// TIA Portal project "V20 Project_V20" (V20)

(* hardware
DEVICE "S7-1500/ET200MP station_1"  S7-1500 station
   slot 0: "Rail_0"  Rack  6ES7 590-1***0-0AA0
   slot 1: "PLC_2"  CPU 1515-2 PN  6ES7 515-2AM00-0AB0  V1.8
      slot 3: "CPU display_1"  6ES7591-1BA00-0AA0
      slot 32768: "PROFINET interface_1"  X1
         slot 32769: "Port_1"  X1 P1
         slot 32770: "Port_2"  X1 P2
      slot 33024: "PROFINET interface_2"  X2
         slot 33025: "Port_1"  X2 P1
*)

// ===== PLC "PLC_2"  CPU 1515-2 PN =====

FUNCTION_BLOCK "FB_CentreStand_Fix_Seq"   // FB1, STL
{ S7_Optimized_Access := 'TRUE' }
VERSION : 0.1
   VAR_INPUT
      iAutoRunning : Bool;
      iFixClamp : Bool;
      iFixEmpty : Bool;
      iFixTrayPresent : Bool;
      iFixUnclamp : Bool;
      iR1DropOver : Bool;
      iR1PickOver : Bool;
      iR2OperationOver : Bool;
      iR2ServiceActivated : Bool;
      iR2ServiceCompleted : Bool;
      iReset_fault : Bool;
      iRobotOutofZone : Bool;
      iSstMode : Bool;
      iSstPB : Bool;
   END_VAR
   VAR_OUTPUT
      qFixClamp : Bool;
      qFixUnclamp : Bool;
      qR1ReadytoDropTray : Bool;
      qR1ReadytoPickTray : Bool;
      qR2OperationStart : Bool;
   END_VAR
   VAR_IN_OUT
      iqR2ServiceActive : Bool;
      iqR2ServiceCompleted : Bool;
   END_VAR
   VAR
      StateNo : Int;
      s138_WaitBothRbtOutAl : Bool;
      s138_WaitBothRbtOutAl_T1 : Bool;
      s138_WaitBothRbtOutAl_T2 : Bool;
      s139_FixEmpty : Bool;
      s139_FixEmpty_T1 : Bool;
      s140_FixTrayPrsntRec : Bool;
      s140_FixTrayPrsntRec_T1 : Bool;
      s140_FixTrayPrsntRec_T2 : Bool;
      s141_FixUnclampCmd : Bool;
      s141_FixUnclampCmd_T1 : Bool;
      s142_TrayRdyDropFix : Bool;
      s142_TrayRdyDropFix_T1 : Bool;
      s143_RbtDropFixChkTr : Bool;
      s143_RbtDropFixChkTr_T1 : Bool;
      s144_RbtOutAreaDrop : Bool;
      s144_RbtOutAreaDrop_T1 : Bool;
      s145_FixClamp : Bool;
      s145_FixClamp_T1 : Bool;
      s146_Rbt2AlloyOpOver : Bool;
      s146_Rbt2AlloyOpOver_T1 : Bool;
      s147_FixUnclmpCmdOvr : Bool;
      s147_FixUnclmpCmdOvr_T1 : Bool;
      s148_RdyPickTrayWait : Bool;
      s148_RdyPickTrayWait_T1 : Bool;
      s149_RbtPickTrayChkEm : Bool;
      s149_RbtPickTrayChkEm_T1 : Bool;
      s191_WaitRbt2OutArea : Bool;
      s191_WaitRbt2OutArea_T1 : Bool;
      sSst : Bool;
      sSstPulse : Bool;
      sSstRise : Bool;
      sStWtResetRel : Bool;
      sStWtResetRel_T1 : Bool;
   END_VAR
   VAR_TEMP
      tOne : Bool;
   END_VAR
BEGIN

REGION Network 1
         O     #tOne;
         ON    #tOne;
         =     #tOne;
END_REGION

REGION Network 2: Create Single Step Pulse bit
         A     #iSstPB;
         FP    #sSstRise;
         =     #sSstPulse;
END_REGION

REGION Network 3: Create Single Step bit
         A     #iSstMode;
         A     #sSstPulse;
         ON    #iSstMode;
         =     #sSst;
END_REGION

REGION Network 4: Transition for STATE Num:0 Reset Released
         A     #sStWtResetRel;
         A     #iAutoRunning;
         =     #sStWtResetRel_T1;
END_REGION

REGION Network 5: STATE Num:0 Reset Released
         A(;
         O     #sStWtResetRel;
         ON    #iAutoRunning;
         );
         AN    #sStWtResetRel_T1;
         =     <??.?>;
         A     <??.?>;
         BLD   102;
         =     #sStWtResetRel;
         A     <??.?>;
         JNB   Label_0;
         L     0;
         T     #StateNo;
   Label_0:NOP   0;
END_REGION

REGION Network 6: Transition for STATE Num:138 Wait for Both Robots Out of Alloy Fixture Center Stand
         A     #s138_WaitBothRbtOutAl;
         AN    #sStWtResetRel;
         A     #sSst;
         =     <??.?>;
         A     <??.?>;
         A     #iRobotOutofZone;
         AN    #iFixTrayPresent;
         =     #s138_WaitBothRbtOutAl_T1;
         A     <??.?>;
         AN    #s138_WaitBothRbtOutAl_T1;
         A     #iRobotOutofZone;
         A     #iFixTrayPresent;
         =     #s138_WaitBothRbtOutAl_T2;
END_REGION

REGION Network 7: STATE Num:138 Wait for Both Robots Out of Alloy Fixture Center Stand
         A(;
         O     #s138_WaitBothRbtOutAl;
         O     #s149_RbtPickTrayChkEm_T1;
         O     #sStWtResetRel_T1;
         );
         AN    #sStWtResetRel;
         AN    #s138_WaitBothRbtOutAl_T1;
         AN    #s138_WaitBothRbtOutAl_T2;
         =     <??.?>;
         A     <??.?>;
         BLD   102;
         =     #s138_WaitBothRbtOutAl;
         A     <??.?>;
         JNB   Label_138;
         L     138;
         T     #StateNo;
   Label_138:NOP   0;
END_REGION

REGION Network 8: Transition for STATE Num:139 Fix Empty
         A     #s139_FixEmpty;
         AN    #sStWtResetRel;
         A     #sSst;
         A     #iFixEmpty;
         =     #s139_FixEmpty_T1;
END_REGION

REGION Network 9: STATE Num:139 Fix Empty
         A(;
         O     #s139_FixEmpty;
         O     #s138_WaitBothRbtOutAl_T1;
         );
         AN    #sStWtResetRel;
         AN    #s139_FixEmpty_T1;
         =     <??.?>;
         A     <??.?>;
         BLD   102;
         =     #s139_FixEmpty;
         A     <??.?>;
         JNB   Label_139;
         L     139;
         T     #StateNo;
   Label_139:NOP   0;
END_REGION

REGION Network 10: Transition for STATE Num:140 Fix Tray Present_Rec Operation pending
         A     #s140_FixTrayPrsntRec;
         AN    #sStWtResetRel;
         A     #sSst;
         =     <??.?>;
         A     <??.?>;
         A     #iFixTrayPresent;
         A     #iRobotOutofZone;
         AN    #iqR2ServiceCompleted;
         =     #s140_FixTrayPrsntRec_T1;
         A     <??.?>;
         AN    #s140_FixTrayPrsntRec_T1;
         A     #iFixTrayPresent;
         A     #iRobotOutofZone;
         A     #iqR2ServiceCompleted;
         =     #s140_FixTrayPrsntRec_T2;
END_REGION

REGION Network 11: STATE Num:140 Fix Tray Present_Rec Operation pending
         A(;
         O     #s140_FixTrayPrsntRec;
         O     #s138_WaitBothRbtOutAl_T2;
         );
         AN    #sStWtResetRel;
         AN    #s140_FixTrayPrsntRec_T1;
         AN    #s140_FixTrayPrsntRec_T2;
         =     <??.?>;
         A     <??.?>;
         BLD   102;
         =     #s140_FixTrayPrsntRec;
         A     <??.?>;
         JNB   Label_140;
         L     140;
         T     #StateNo;
   Label_140:NOP   0;
END_REGION

REGION Network 12: Transition for STATE Num:141 Fix Unclamp Cmd
         A     #s141_FixUnclampCmd;
         AN    #sStWtResetRel;
         A     #sSst;
         A     #iFixUnclamp;
         =     #s141_FixUnclampCmd_T1;
END_REGION

REGION Network 13: STATE Num:141 Fix Unclamp Cmd
         A(;
         O     #s141_FixUnclampCmd;
         O     #s139_FixEmpty_T1;
         );
         AN    #sStWtResetRel;
         AN    #s141_FixUnclampCmd_T1;
         =     <??.?>;
         A     <??.?>;
         BLD   102;
         =     #s141_FixUnclampCmd;
         A     <??.?>;
         JNB   Label_141;
         L     141;
         T     #StateNo;
   Label_141:NOP   0;
END_REGION

REGION Network 14: Actions for STATE Num:141 Fix Unclamp Cmd
         A     #s141_FixUnclampCmd;
         =     #qFixUnclamp;
END_REGION

REGION Network 15: Transition for STATE Num:142 Tray Rdy to Drop Fix- Wait for Robot Accept request
         A     #s142_TrayRdyDropFix;
         AN    #sStWtResetRel;
         A     #sSst;
         A     #iR1DropOver;
         =     #s142_TrayRdyDropFix_T1;
END_REGION

REGION Network 16: STATE Num:142 Tray Rdy to Drop Fix- Wait for Robot Accept request
         A(;
         O     #s142_TrayRdyDropFix;
         O     #s141_FixUnclampCmd_T1;
         );
         AN    #sStWtResetRel;
         AN    #s142_TrayRdyDropFix_T1;
         =     <??.?>;
         A     <??.?>;
         BLD   102;
         =     #s142_TrayRdyDropFix;
         A     <??.?>;
         JNB   Label_142;
         L     142;
         T     #StateNo;
   Label_142:NOP   0;
END_REGION

REGION Network 17: Actions for STATE Num:142 Tray Rdy to Drop Fix- Wait for Robot Accept request
         A     #s142_TrayRdyDropFix;
         =     #qR1ReadytoDropTray;
END_REGION

REGION Network 18: Transition for STATE Num:143 Robot Drop Fix and Check Tray Present
         A     #s143_RbtDropFixChkTr;
         AN    #sStWtResetRel;
         A     #sSst;
         A     #iFixTrayPresent;
         =     #s143_RbtDropFixChkTr_T1;
END_REGION

REGION Network 19: STATE Num:143 Robot Drop Fix and Check Tray Present
         A(;
         O     #s143_RbtDropFixChkTr;
         O     #s142_TrayRdyDropFix_T1;
         );
         AN    #sStWtResetRel;
         AN    #s143_RbtDropFixChkTr_T1;
         =     <??.?>;
         A     <??.?>;
         BLD   102;
         =     #s143_RbtDropFixChkTr;
         A     <??.?>;
         JNB   Label_143;
         L     143;
         T     #StateNo;
   Label_143:NOP   0;
END_REGION

REGION Network 20: Transition for STATE Num:144 Rbt Out of Area After Drop
         A     #s144_RbtOutAreaDrop;
         AN    #sStWtResetRel;
         A     #sSst;
         A     #iRobotOutofZone;
         =     #s144_RbtOutAreaDrop_T1;
END_REGION

REGION Network 21: STATE Num:144 Rbt Out of Area After Drop
         A(;
         O     #s144_RbtOutAreaDrop;
         O     #s143_RbtDropFixChkTr_T1;
         );
         AN    #sStWtResetRel;
         AN    #s144_RbtOutAreaDrop_T1;
         =     <??.?>;
         A     <??.?>;
         BLD   102;
         =     #s144_RbtOutAreaDrop;
         A     <??.?>;
         JNB   Label_144;
         L     144;
         T     #StateNo;
   Label_144:NOP   0;
END_REGION

REGION Network 22: Transition for STATE Num:145 Fix Clamp
         A     #s145_FixClamp;
         AN    #sStWtResetRel;
         A     #sSst;
         A     #iRobotOutofZone;
         A     #iFixClamp;
         =     #s145_FixClamp_T1;
END_REGION

REGION Network 23: STATE Num:145 Fix Clamp
         A(;
         O     #s145_FixClamp;
         O     #s140_FixTrayPrsntRec_T1;
         O     #s144_RbtOutAreaDrop_T1;
         );
         AN    #sStWtResetRel;
         AN    #s145_FixClamp_T1;
         =     <??.?>;
         A     <??.?>;
         BLD   102;
         =     #s145_FixClamp;
         A     <??.?>;
         JNB   Label_145;
         L     145;
         T     #StateNo;
   Label_145:NOP   0;
END_REGION

REGION Network 24: Actions for STATE Num:145 Fix Clamp
         A     #s145_FixClamp;
         =     #qFixClamp;
END_REGION

REGION Network 25: Transition for STATE Num:146 Robot-2 All Alloys Pick Or Drop Operation over
         A     #s146_Rbt2AlloyOpOver;
         AN    #sStWtResetRel;
         A     #sSst;
         A     #iR2OperationOver;
         =     #s146_Rbt2AlloyOpOver_T1;
END_REGION

REGION Network 26: STATE Num:146 Robot-2 All Alloys Pick Or Drop Operation over
         A(;
         O     #s146_Rbt2AlloyOpOver;
         O     #s145_FixClamp_T1;
         );
         AN    #sStWtResetRel;
         AN    #s146_Rbt2AlloyOpOver_T1;
         =     <??.?>;
         A     <??.?>;
         BLD   102;
         =     #s146_Rbt2AlloyOpOver;
         A     <??.?>;
         JNB   Label_146;
         L     146;
         T     #StateNo;
   Label_146:NOP   0;
END_REGION

REGION Network 27: Actions for STATE Num:146 Robot-2 All Alloys Pick Or Drop Operation over
         A     #s146_Rbt2AlloyOpOver;
         =     #qR2OperationStart;
         A     #iR2ServiceActivated;
         S     #iqR2ServiceActive;
         A     #iR2OperationOver;
         A     #iqR2ServiceActive;
         R     #iqR2ServiceActive;
END_REGION

REGION Network 28: Transition for STATE Num:147 Fix Unclamp Cmd After Opern over
         A     #s147_FixUnclmpCmdOvr;
         AN    #sStWtResetRel;
         A     #sSst;
         A     #iFixUnclamp;
         =     #s147_FixUnclmpCmdOvr_T1;
END_REGION

REGION Network 29: STATE Num:147 Fix Unclamp Cmd After Opern over
         A(;
         O     #s147_FixUnclmpCmdOvr;
         O     #s140_FixTrayPrsntRec_T2;
         O     #s191_WaitRbt2OutArea_T1;
         );
         AN    #sStWtResetRel;
         AN    #s147_FixUnclmpCmdOvr_T1;
         =     <??.?>;
         A     <??.?>;
         BLD   102;
         =     #s147_FixUnclmpCmdOvr;
         A     <??.?>;
         JNB   Label_147;
         L     147;
         T     #StateNo;
   Label_147:NOP   0;
END_REGION

REGION Network 30: Actions for STATE Num:147 Fix Unclamp Cmd After Opern over
         A     #s147_FixUnclmpCmdOvr;
         =     #qFixUnclamp;
END_REGION

REGION Network 31: Transition for STATE Num:148 Rdy to Pick Tray After Oprn Over- Wait for Robot Accept Request
         A     #s148_RdyPickTrayWait;
         AN    #sStWtResetRel;
         A     #sSst;
         A     #iR1PickOver;
         =     #s148_RdyPickTrayWait_T1;
END_REGION

REGION Network 32: STATE Num:148 Rdy to Pick Tray After Oprn Over- Wait for Robot Accept Request
         A(;
         O     #s148_RdyPickTrayWait;
         O     #s147_FixUnclmpCmdOvr_T1;
         );
         AN    #sStWtResetRel;
         AN    #s148_RdyPickTrayWait_T1;
         =     <??.?>;
         A     <??.?>;
         BLD   102;
         =     #s148_RdyPickTrayWait;
         A     <??.?>;
         JNB   Label_148;
         L     148;
         T     #StateNo;
   Label_148:NOP   0;
END_REGION

REGION Network 33: Actions for STATE Num:148 Rdy to Pick Tray After Oprn Over- Wait for Robot Accept Request
         A     #s148_RdyPickTrayWait;
         =     #qR1ReadytoPickTray;
         A     #iR1PickOver;
         R     #iqR2ServiceCompleted;
END_REGION

REGION Network 34: Transition for STATE Num:149 Robot Picked Tray and Check Tray Loc Empty
         A     #s149_RbtPickTrayChkEm;
         AN    #sStWtResetRel;
         A     #sSst;
         A     #iFixEmpty;
         =     #s149_RbtPickTrayChkEm_T1;
END_REGION

REGION Network 35: STATE Num:149 Robot Picked Tray and Check Tray Loc Empty
         A(;
         O     #s149_RbtPickTrayChkEm;
         O     #s148_RdyPickTrayWait_T1;
         );
         AN    #sStWtResetRel;
         AN    #s149_RbtPickTrayChkEm_T1;
         =     <??.?>;
         A     <??.?>;
         BLD   102;
         =     #s149_RbtPickTrayChkEm;
         A     <??.?>;
         JNB   Label_149;
         L     149;
         T     #StateNo;
   Label_149:NOP   0;
END_REGION

REGION Network 36: Actions for STATE Num:149 Robot Picked Tray and Check Tray Loc Empty
         A     #s149_RbtPickTrayChkEm;
         R     #iqR2ServiceCompleted;
END_REGION

REGION Network 37: Transition for STATE Num:191 Wait For Robot-2 Out Of Area
         A     #s191_WaitRbt2OutArea;
         AN    #sStWtResetRel;
         A     #sSst;
         A     #iRobotOutofZone;
         =     #s191_WaitRbt2OutArea_T1;
END_REGION

REGION Network 38: STATE Num:191 Wait For Robot-2 Out Of Area
         A(;
         O     #s191_WaitRbt2OutArea;
         O     #s146_Rbt2AlloyOpOver_T1;
         );
         AN    #sStWtResetRel;
         AN    #s191_WaitRbt2OutArea_T1;
         =     <??.?>;
         A     <??.?>;
         BLD   102;
         =     #s191_WaitRbt2OutArea;
         A     <??.?>;
         JNB   Label_191;
         L     191;
         T     #StateNo;
   Label_191:NOP   0;
END_REGION
END_FUNCTION_BLOCK

FUNCTION_BLOCK "Block_1"   // FB1, LAD
{ S7_Optimized_Access := 'TRUE' }
BEGIN

REGION Network 1
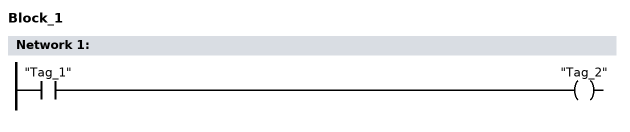
   RUNG wire#powerrail
      Contact( "Tag_1" )
      Coil( "Tag_2" )
   END_RUNG
   // the same network as SCL:
   "Tag_2" := "Tag_1";
END_REGION
END_FUNCTION_BLOCK

ORGANIZATION_BLOCK "Main"   // OB1, LAD, ProgramCycle
TITLE = "Main Program Sweep (Cycle)"
{ S7_Optimized_Access := 'TRUE' }
VERSION : 0.1
   VAR_INPUT
      Initial_Call : Bool;   // Initial call of this OB
      Remanence : Bool;   // =True, if remanent data are available
   END_VAR
BEGIN
END_ORGANIZATION_BLOCK

// ===== library types =====

// folder: SM-Modules

FUNCTION_BLOCK "PR_TT3PosControl"   // FB335, LAD
TITLE = PR_TT3PosControl
{ S7_Optimized_Access := 'TRUE' }
AUTHOR : Virendra Sharma
FAMILY : Wipro_Pari
NAME : SM0106022020
VERSION : 0.1
   VAR_INPUT
      iResetFaults : Bool;   // Reset Fault input
      iControlOn : Bool;   // Control On Input
      iPos1Cmd : Bool;   // Zero degree position command (Home position)
      iPos2Cmd : Bool;   // Plus 90 degree position command
      iPos3Cmd : Bool;   // Minus 90 degree position command
      iPos1StopSens : Bool;   // zero degree position stop sensor
      iPos2StopSens : Bool;   // Plus 90 degree position stop sensor
      iPos3StopSens : Bool;   // Minus 90 degree position stop sensor
      iTimeForPosOver : Time;   // Timer Value for position over
      iTimeForVFDStop : Time;   // Time value for VFD stop
      iPositiveOTLS : Bool;   // Positive direction over travel limit swithch
      iNegativeOTLS : Bool;   // Negative direction over travel limit swithch
      iFwdInterlock : Bool;   // Connect Forward Interlock Conditions
      iRevInterlock : Bool;   // Connect Reverse Interlock Conditions
      iVFDRunning : Bool;
   END_VAR
   VAR_OUTPUT
      qPos1Over : Bool;   // Zero position over
      qPos2Over : Bool;   // Plus 90 position
      qPos3Over : Bool;   // Minus 90 position over
      qVFDFwd : Bool;   // VFD Rotating Forward
      qVFDRev : Bool;   // VFD Rotating Reverse
      qModuleFault : Bool;   // Error Module Fault
      qError : Array[0..7] of Bool;   // Error Forward Interlock
      qMsg : Array[0..7] of Bool;
   END_VAR
   VAR
      sFaultReset : Bool;
      sFwdCmdOn : Bool;
      sDriveRdyFrCmd : Bool;
      sTimeForPosOver : Time;
      sTimeForVFDStop : Time;
      sRevCmdOn : Bool;
      sCtrlFrmNet : Bool;
      sRefFrmNet : Bool;
      sTimerOn : Bool;
      s0PosCmdActive : Bool;
      s0PosActiveForFwd : Bool;
      s0PosActiveForRev : Bool;
      s0PosActiveForFwdOver : Bool;
      s0PosActiveForRevOver : Bool;
      s0PosOverTON : TON_TIME;
      sMinus90PosActiveForRev : Bool;
      sMinus90PosCmdActive : Bool;
      sMinus90PosOverTON : TON_TIME;
      sMinus90PosActiveForFwdOver : Bool;
      sMinus90PosActiveForRevOver : Bool;
      sPlus90PosActiveForFwd : Bool;
      sPlus90PosCmdActive : Bool;
      sPlus90PosOverTON : TON_TIME;
      sPlus90PosActiveForFwdOver : Bool;
      sPlus90PosActiveForRevOver : Bool;
      sTTAtPos0 : Bool;
      sTTAtPos0Done : Bool;
      sTTAtPosMinus90 : Bool;
      sTTAtPosMinus90Done : Bool;
      sTTAtPosPlus90 : Bool;
      sTTAtPosPlus90Done : Bool;
      sPuls : Array[0..16] of Bool;
   END_VAR
   VAR RETAIN
      sTargetPos : Word;
      sLastPos : Word;
   END_VAR
   VAR
      sVFDFwdRunning : Bool;
      sVFDRunningDlyDn : TON_TIME;
      sVFDRevRunning : Bool;
      sFwdInterlockErr : Bool;
      sRevInterlockErr : Bool;
      sPositiveOTLSErr : Bool;
      sNegativeOTLSErr : Bool;
      sVFDStopped : Bool;
   END_VAR
   VAR RETAIN
      sFwdActiveFor1ToPos2 : Bool;
      sRevAvtiveFor1ToPos3 : Bool;
      sFwdActiveFor3ToPos1 : Bool;
      sRevAvtiveFor2ToPos1 : Bool;
   END_VAR
   VAR_TEMP   // added for the SCL form of the ladder/FBD networks
      _w1 : Bool;
      _w2 : Bool;
      _w3 : Bool;
      _w4 : Bool;
      _w5 : Bool;
      _w6 : Bool;
   END_VAR
   // // qError[1] : Error Reverse Interlock
   // // qError[2] : Error Forward Interlock
   // // qError[3] : Turn Table over traveled at positive side
   // // qError[4] : Turn Table over traveled at negative side
   // // qError[0] : Error VFD Stopped
   // // qMsg[0] : TT not referenced.
BEGIN

REGION Network 1: Header
   // ==============================================================================
   //  Company: Precision Automation & Robotics India Ltd. (WIPRO-PARI)
   // ------------------------------------------------------------------------------
   //  Item Code: SM0106022020
   //  Author/Created by: Virendra Sharma
   //  Reviewed/Checked by: Sandip Chavanke
   //  First Release on: 11-Oct-2023
   //  Latest update on: 11-Oct-2023
   // ------------------------------------------------------------------------------
   //  Tested with: CPU firmware, model or simulator testing
   //  Engineering/Editor: TIA Portal V17
   // ------------------------------------------------------------------------------
   //  Restrictions: More then 3 Position of turn table
   //  Dependencies/Requirements:
   //  <hardware, technology package, memory needed, data types (UDT's), other blocks, etc.>
   // ------------------------------------------------------------------------------
   //  Change Log:
   //  Ver.	Date		Changed by		Details of changes
   //  1.0	11-10-2023	Virendra Sharma 	First release version- 1.0
   // ------------------------------------------------------------------------------
   //  Functionality: This Module is to control the motion of VFD that controls Turn Table with 3 distinctive positions,
   //  like home or Path1 (0 Degree), Path3 (Minus 90 Degree), and path2 (Plus 90 Degree) positions.
   //  Each position is provided with a 'position sensor' to confirm the position of the Turn Table and to stop the Turn Table at the given position.
   //  The position of the turn table is defined by where the main stopper is located.
   //  <include block inputs, outputs, in-outs>
   //  Inputs
   //  1. iResetFaults : Bool
   //  2. iControlOn : Bool
   //  3. iPos1Cmd : Bool
   //  4. iPos2Cmd : Bool
   //  5. iPos3Cmd : Bool
   //  6. iPos1StopSens : Bool
   //  7. iPos2StopSens : Bool
   //  8. iPos3StopSens : Bool
   //  9. iTimeForPosOver : Time
   //  10. iTimeForVFDStop : Time
   //  11. iPositiveOTLS : Bool
   //  12. iNegativeOTLS : Bool
   //  13. iFwdInterlock : Bool
   //  14. iRevInterlock : Bool
   // 
   //  Outputs
   //  1. qPos1Over : Bool
   //  2. qPos2Over : Bool
   //  3. qPos3Over : Bool
   //  4. qVFDFwd : Bool
   //  5. qVFDRev : Bool
   //  6. qModuleFault : bool
   //  7. qError : Array [0..31] of Bool
   //  8. qMsg : Array [0..31] of Bool  
   // 
   //  In-outs
   //  NA
   // ------------------------------------------------------------------------------
   //  Errors reported:
   //  1. Error 0 : Error VFD Stopped
   //  2. Error 1 : Error Reverse Interlock 
   //  3. Error 2 : Error Forward Interlock 
   //  4. Error 3 : Turn Table over traveled at positive side
   //  5. Error 4 : Turn Table over traveled at negative side
   //  Messages reported:
   //  1. Message 0 : TT not referenced.
   // ==============================================================================
END_REGION

REGION Network 2: Fault Reset
   // Error reset request flag
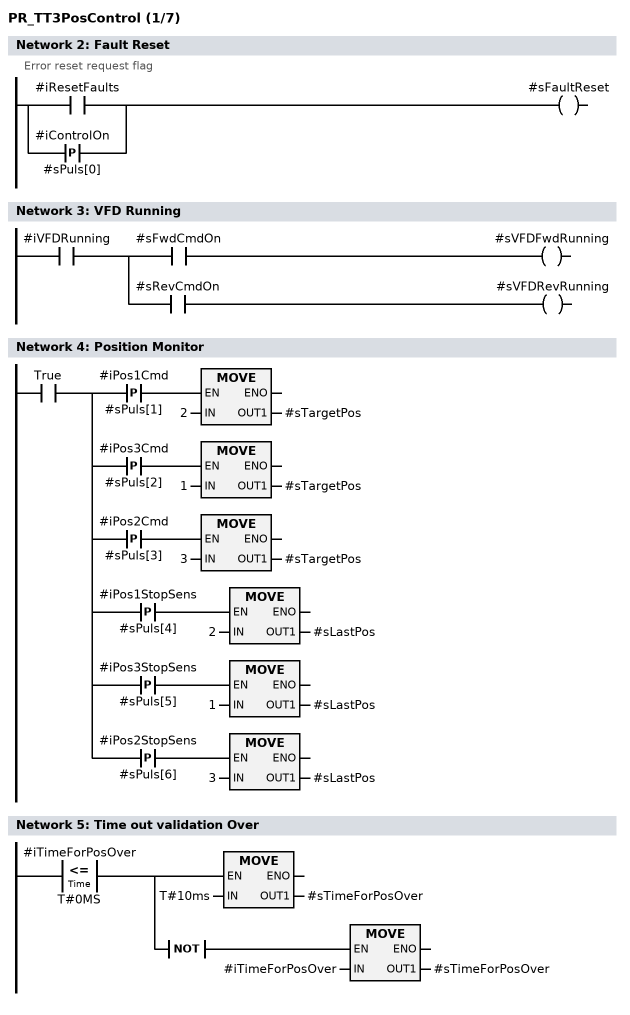
   RUNG wire#powerrail
      Contact( #iResetFaults )
      wire#w1
      Coil( #sFaultReset )
   END_RUNG
   RUNG wire#powerrail
      P_Contact(operand := #iControlOn, bit := #sPuls[0])
   END_RUNG wire#w1
   // the same network as SCL:
   #_w1 := #iControlOn AND NOT #sPuls[0];   // rising edge of #iControlOn
   #sPuls[0] := #iControlOn;
   #sFaultReset := #iResetFaults OR #_w1;
END_REGION

REGION Network 3: VFD Running
   RUNG wire#powerrail
      Contact( #iVFDRunning )
      wire#w1
      Contact( #sFwdCmdOn )
      Coil( #sVFDFwdRunning )
   END_RUNG
   RUNG wire#w1
      Contact( #sRevCmdOn )
      Coil( #sVFDRevRunning )
   END_RUNG
   // the same network as SCL:
   #sVFDFwdRunning := #iVFDRunning AND #sFwdCmdOn;
   #sVFDRevRunning := #iVFDRunning AND #sRevCmdOn;
END_REGION

REGION Network 4: Position Monitor
   RUNG wire#powerrail
      Contact( True )
      wire#w1
      P_Contact(operand := #iPos1Cmd, bit := #sPuls[1])
      Move(in := 2, out1 => #sTargetPos)
   END_RUNG
   RUNG wire#w1
      P_Contact(operand := #iPos3Cmd, bit := #sPuls[2])
      Move(in := 1, out1 => #sTargetPos)
   END_RUNG
   RUNG wire#w1
      P_Contact(operand := #iPos2Cmd, bit := #sPuls[3])
      Move(in := 3, out1 => #sTargetPos)
   END_RUNG
   RUNG wire#w1
      P_Contact(operand := #iPos1StopSens, bit := #sPuls[4])
      Move(in := 2, out1 => #sLastPos)
   END_RUNG
   RUNG wire#w1
      P_Contact(operand := #iPos3StopSens, bit := #sPuls[5])
      Move(in := 1, out1 => #sLastPos)
   END_RUNG
   RUNG wire#w1
      P_Contact(operand := #iPos2StopSens, bit := #sPuls[6])
      Move(in := 3, out1 => #sLastPos)
   END_RUNG
   // the same network as SCL:
   #_w1 := True AND #iPos1Cmd AND NOT #sPuls[1];   // rising edge of #iPos1Cmd
   #sPuls[1] := #iPos1Cmd;
   IF #_w1 THEN #sTargetPos := 2; END_IF;
   #_w2 := True AND #iPos3Cmd AND NOT #sPuls[2];   // rising edge of #iPos3Cmd
   #sPuls[2] := #iPos3Cmd;
   IF #_w2 THEN #sTargetPos := 1; END_IF;
   #_w3 := True AND #iPos2Cmd AND NOT #sPuls[3];   // rising edge of #iPos2Cmd
   #sPuls[3] := #iPos2Cmd;
   IF #_w3 THEN #sTargetPos := 3; END_IF;
   #_w4 := True AND #iPos1StopSens AND NOT #sPuls[4];   // rising edge of #iPos1StopSens
   #sPuls[4] := #iPos1StopSens;
   IF #_w4 THEN #sLastPos := 2; END_IF;
   #_w5 := True AND #iPos3StopSens AND NOT #sPuls[5];   // rising edge of #iPos3StopSens
   #sPuls[5] := #iPos3StopSens;
   IF #_w5 THEN #sLastPos := 1; END_IF;
   #_w6 := True AND #iPos2StopSens AND NOT #sPuls[6];   // rising edge of #iPos2StopSens
   #sPuls[6] := #iPos2StopSens;
   IF #_w6 THEN #sLastPos := 3; END_IF;
END_REGION

REGION Network 5: Time out validation Over
   RUNG wire#powerrail
      { S7_Templates := "SrcType := Time" } LE_Contact(in1 := #iTimeForPosOver, in2 := T#0MS)
      wire#w1
      Move(in := T#10ms, out1 => #sTimeForPosOver)
   END_RUNG
   RUNG wire#w1
      Not()
      Move(in := #iTimeForPosOver, out1 => #sTimeForPosOver)
   END_RUNG
   // the same network as SCL:
   #_w1 := #iTimeForPosOver <= T#0MS;
   IF #_w1 THEN #sTimeForPosOver := T#10ms; END_IF;
   IF NOT #_w1 THEN #sTimeForPosOver := #iTimeForPosOver; END_IF;
END_REGION

REGION Network 6: In Zone command form Positon 1
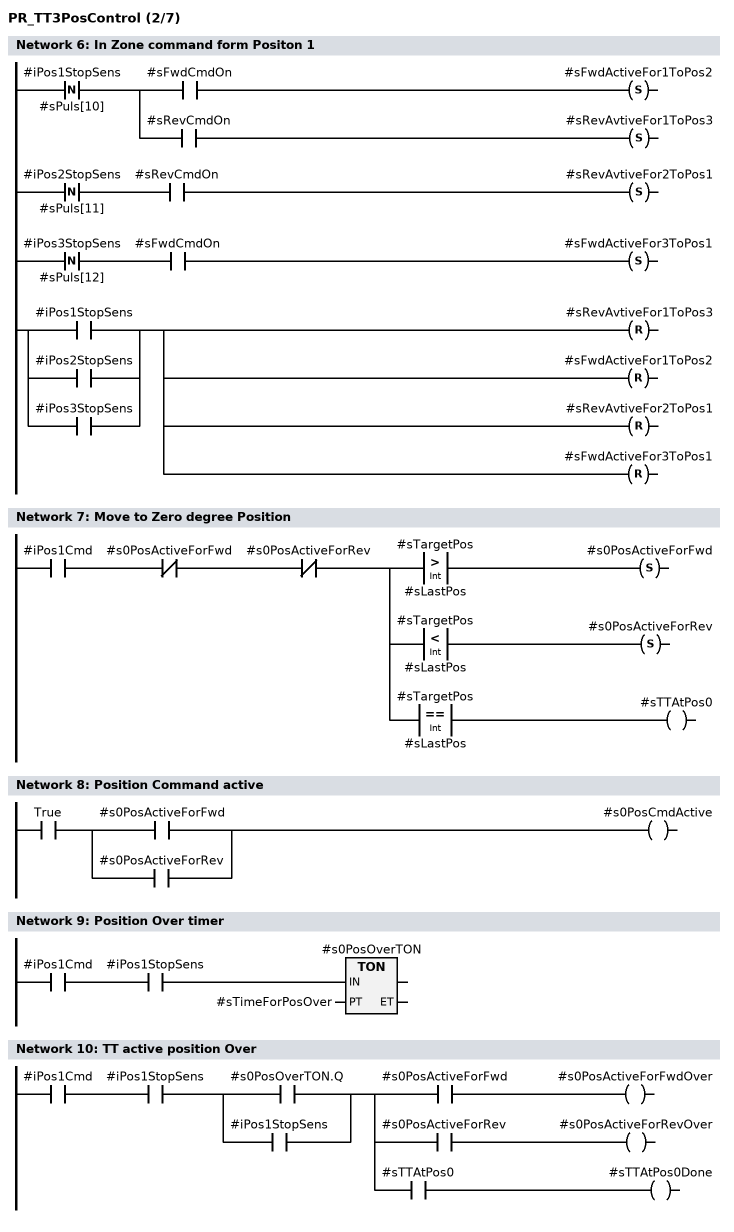
   RUNG wire#powerrail
      N_Contact(operand := #iPos1StopSens, bit := #sPuls[10])
      wire#w1
      Contact( #sFwdCmdOn )
      S_Coil( #sFwdActiveFor1ToPos2 )
   END_RUNG
   RUNG wire#w1
      Contact( #sRevCmdOn )
      S_Coil( #sRevAvtiveFor1ToPos3 )
   END_RUNG
   RUNG wire#powerrail
      N_Contact(operand := #iPos2StopSens, bit := #sPuls[11])
      Contact( #sRevCmdOn )
      S_Coil( #sRevAvtiveFor2ToPos1 )
   END_RUNG
   RUNG wire#powerrail
      N_Contact(operand := #iPos3StopSens, bit := #sPuls[12])
      Contact( #sFwdCmdOn )
      S_Coil( #sFwdActiveFor3ToPos1 )
   END_RUNG
   RUNG wire#powerrail
      Contact( #iPos1StopSens )
      wire#w2
      R_Coil( #sRevAvtiveFor1ToPos3 )
   END_RUNG
   RUNG wire#powerrail
      Contact( #iPos2StopSens )
   END_RUNG wire#w2
   RUNG wire#powerrail
      Contact( #iPos3StopSens )
   END_RUNG wire#w2
   RUNG wire#w2
      R_Coil( #sFwdActiveFor1ToPos2 )
   END_RUNG
   RUNG wire#w2
      R_Coil( #sRevAvtiveFor2ToPos1 )
   END_RUNG
   RUNG wire#w2
      R_Coil( #sFwdActiveFor3ToPos1 )
   END_RUNG
   // the same network as SCL:
   #_w1 := NOT #iPos1StopSens AND #sPuls[10];   // falling edge of #iPos1StopSens
   #sPuls[10] := #iPos1StopSens;
   IF #_w1 AND #sFwdCmdOn THEN #sFwdActiveFor1ToPos2 := TRUE; END_IF;
   IF #_w1 AND #sRevCmdOn THEN #sRevAvtiveFor1ToPos3 := TRUE; END_IF;
   #_w2 := NOT #iPos2StopSens AND #sPuls[11];   // falling edge of #iPos2StopSens
   #sPuls[11] := #iPos2StopSens;
   IF #_w2 AND #sRevCmdOn THEN #sRevAvtiveFor2ToPos1 := TRUE; END_IF;
   #_w3 := NOT #iPos3StopSens AND #sPuls[12];   // falling edge of #iPos3StopSens
   #sPuls[12] := #iPos3StopSens;
   IF #_w3 AND #sFwdCmdOn THEN #sFwdActiveFor3ToPos1 := TRUE; END_IF;
   IF #iPos1StopSens OR #iPos2StopSens OR #iPos3StopSens THEN
       #sRevAvtiveFor1ToPos3 := FALSE;
       #sFwdActiveFor1ToPos2 := FALSE;
       #sRevAvtiveFor2ToPos1 := FALSE;
       #sFwdActiveFor3ToPos1 := FALSE;
   END_IF;
END_REGION

REGION Network 7: Move to Zero degree Position
   RUNG wire#powerrail
      Contact( #iPos1Cmd )
      I_Contact( #s0PosActiveForFwd )
      I_Contact( #s0PosActiveForRev )
      wire#w1
      { S7_Templates := "SrcType := Int" } GT_Contact(in1 := #sTargetPos, in2 := #sLastPos)
      S_Coil( #s0PosActiveForFwd )
   END_RUNG
   RUNG wire#w1
      { S7_Templates := "SrcType := Int" } LT_Contact(in1 := #sTargetPos, in2 := #sLastPos)
      S_Coil( #s0PosActiveForRev )
   END_RUNG
   RUNG wire#w1
      { S7_Templates := "SrcType := Int" } EQ_Contact(in1 := #sTargetPos, in2 := #sLastPos)
      Coil( #sTTAtPos0 )
   END_RUNG
   // the same network as SCL:
   #_w1 := #iPos1Cmd AND NOT #s0PosActiveForFwd AND NOT #s0PosActiveForRev;
   IF #_w1 AND (#sTargetPos > #sLastPos) THEN #s0PosActiveForFwd := TRUE; END_IF;
   IF #_w1 AND (#sTargetPos < #sLastPos) THEN #s0PosActiveForRev := TRUE; END_IF;
   #sTTAtPos0 := #_w1 AND (#sTargetPos = #sLastPos);
END_REGION

REGION Network 8: Position Command active
   RUNG wire#powerrail
      Contact( True )
      wire#w1
      Contact( #s0PosActiveForFwd )
      wire#w2
      Coil( #s0PosCmdActive )
   END_RUNG
   RUNG wire#w1
      Contact( #s0PosActiveForRev )
   END_RUNG wire#w2
   // the same network as SCL:
   #s0PosCmdActive := True AND (#s0PosActiveForFwd OR #s0PosActiveForRev);
END_REGION

REGION Network 9: Position Over timer
   #s0PosOverTON(IN := #iPos1Cmd AND #iPos1StopSens, PT := #sTimeForPosOver);   // TON
END_REGION

REGION Network 10: TT active position Over
   RUNG wire#powerrail
      Contact( #iPos1Cmd )
      Contact( #iPos1StopSens )
      wire#w1
      Contact( #s0PosOverTON.Q )
      wire#w2
      Contact( #s0PosActiveForFwd )
      Coil( #s0PosActiveForFwdOver )
   END_RUNG
   RUNG wire#w1
      Contact( #iPos1StopSens )
   END_RUNG wire#w2
   RUNG wire#w2
      Contact( #s0PosActiveForRev )
      Coil( #s0PosActiveForRevOver )
   END_RUNG
   RUNG wire#w2
      Contact( #sTTAtPos0 )
      Coil( #sTTAtPos0Done )
   END_RUNG
   // the same network as SCL:
   #_w1 := #iPos1Cmd AND #iPos1StopSens AND (#s0PosOverTON.Q OR #iPos1StopSens);
   #s0PosActiveForFwdOver := #_w1 AND #s0PosActiveForFwd;
   #s0PosActiveForRevOver := #_w1 AND #s0PosActiveForRev;
   #sTTAtPos0Done := #_w1 AND #sTTAtPos0;
END_REGION

REGION Network 11: Position over output
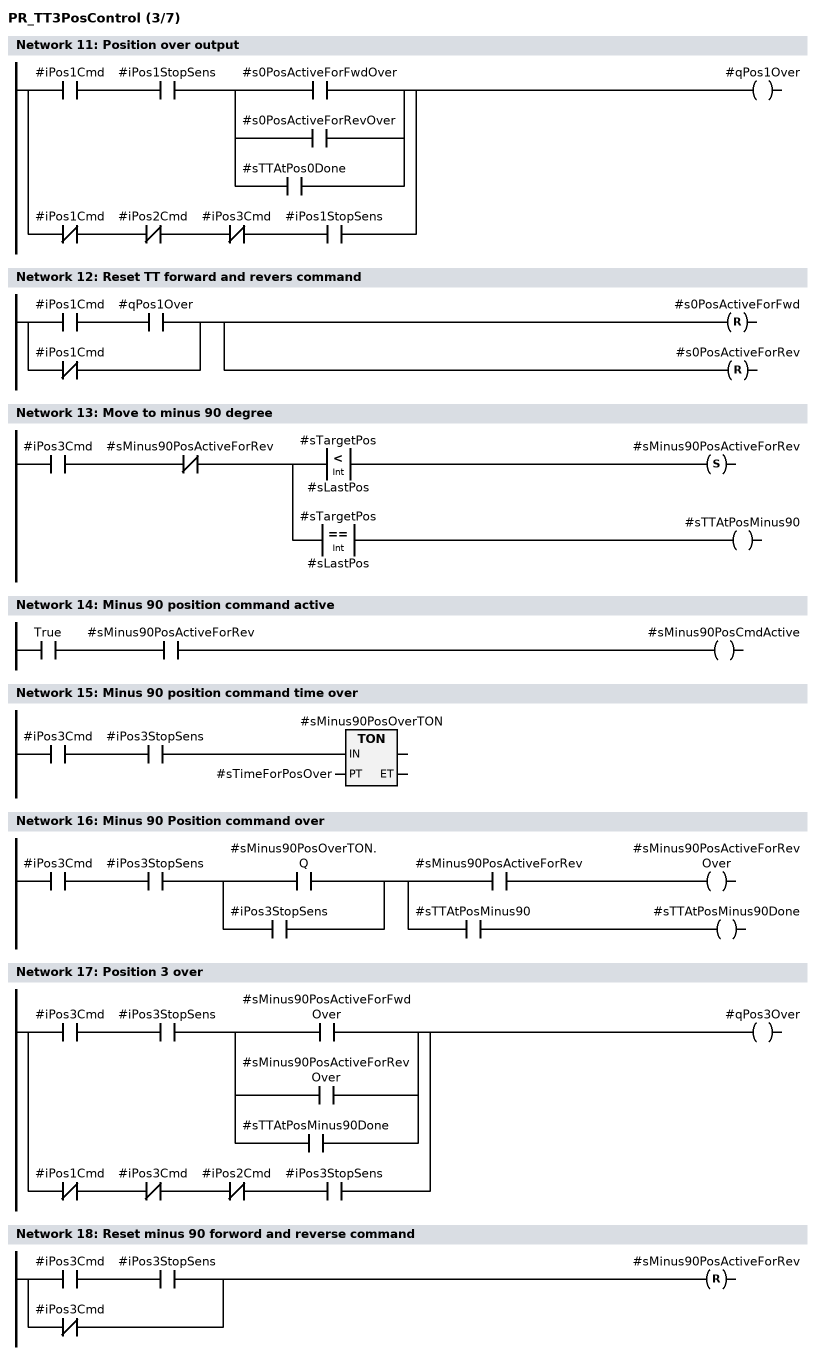
   RUNG wire#powerrail
      Contact( #iPos1Cmd )
      Contact( #iPos1StopSens )
      wire#w1
      Contact( #s0PosActiveForFwdOver )
      wire#w2
      Coil( #qPos1Over )
   END_RUNG
   RUNG wire#w1
      Contact( #s0PosActiveForRevOver )
   END_RUNG wire#w2
   RUNG wire#w1
      Contact( #sTTAtPos0Done )
   END_RUNG wire#w2
   RUNG wire#powerrail
      I_Contact( #iPos1Cmd )
      I_Contact( #iPos2Cmd )
      I_Contact( #iPos3Cmd )
      Contact( #iPos1StopSens )
   END_RUNG wire#w2
   // the same network as SCL:
   #qPos1Over := (#iPos1Cmd AND #iPos1StopSens AND (#s0PosActiveForFwdOver OR #s0PosActiveForRevOver OR #sTTAtPos0Done)) OR (NOT #iPos1Cmd AND NOT #iPos2Cmd AND NOT #iPos3Cmd AND #iPos1StopSens);
END_REGION

REGION Network 12: Reset TT forward and revers command
   RUNG wire#powerrail
      Contact( #iPos1Cmd )
      Contact( #qPos1Over )
      wire#w1
      R_Coil( #s0PosActiveForFwd )
   END_RUNG
   RUNG wire#powerrail
      I_Contact( #iPos1Cmd )
   END_RUNG wire#w1
   RUNG wire#w1
      R_Coil( #s0PosActiveForRev )
   END_RUNG
   // the same network as SCL:
   IF (#iPos1Cmd AND #qPos1Over) OR NOT #iPos1Cmd THEN
       #s0PosActiveForFwd := FALSE;
       #s0PosActiveForRev := FALSE;
   END_IF;
END_REGION

REGION Network 13: Move to minus 90 degree
   RUNG wire#powerrail
      Contact( #iPos3Cmd )
      I_Contact( #sMinus90PosActiveForRev )
      wire#w1
      { S7_Templates := "SrcType := Int" } LT_Contact(in1 := #sTargetPos, in2 := #sLastPos)
      S_Coil( #sMinus90PosActiveForRev )
   END_RUNG
   RUNG wire#w1
      { S7_Templates := "SrcType := Int" } EQ_Contact(in1 := #sTargetPos, in2 := #sLastPos)
      Coil( #sTTAtPosMinus90 )
   END_RUNG
   // the same network as SCL:
   #_w1 := #iPos3Cmd AND NOT #sMinus90PosActiveForRev;
   IF #_w1 AND (#sTargetPos < #sLastPos) THEN #sMinus90PosActiveForRev := TRUE; END_IF;
   #sTTAtPosMinus90 := #_w1 AND (#sTargetPos = #sLastPos);
END_REGION

REGION Network 14: Minus 90 position command active
   RUNG wire#powerrail
      Contact( True )
      Contact( #sMinus90PosActiveForRev )
      Coil( #sMinus90PosCmdActive )
   END_RUNG
   // the same network as SCL:
   #sMinus90PosCmdActive := True AND #sMinus90PosActiveForRev;
END_REGION

REGION Network 15: Minus 90 position command time over
   #sMinus90PosOverTON(IN := #iPos3Cmd AND #iPos3StopSens, PT := #sTimeForPosOver);   // TON
END_REGION

REGION Network 16: Minus 90 Position command over
   RUNG wire#powerrail
      Contact( #iPos3Cmd )
      Contact( #iPos3StopSens )
      wire#w1
      Contact( #sMinus90PosOverTON.Q )
      wire#w2
      Contact( #sMinus90PosActiveForRev )
      Coil( #sMinus90PosActiveForRevOver )
   END_RUNG
   RUNG wire#w1
      Contact( #iPos3StopSens )
   END_RUNG wire#w2
   RUNG wire#w2
      Contact( #sTTAtPosMinus90 )
      Coil( #sTTAtPosMinus90Done )
   END_RUNG
   // the same network as SCL:
   #_w1 := #iPos3Cmd AND #iPos3StopSens AND (#sMinus90PosOverTON.Q OR #iPos3StopSens);
   #sMinus90PosActiveForRevOver := #_w1 AND #sMinus90PosActiveForRev;
   #sTTAtPosMinus90Done := #_w1 AND #sTTAtPosMinus90;
END_REGION

REGION Network 17: Position 3 over
   RUNG wire#powerrail
      Contact( #iPos3Cmd )
      Contact( #iPos3StopSens )
      wire#w1
      Contact( #sMinus90PosActiveForFwdOver )
      wire#w2
      Coil( #qPos3Over )
   END_RUNG
   RUNG wire#w1
      Contact( #sMinus90PosActiveForRevOver )
   END_RUNG wire#w2
   RUNG wire#w1
      Contact( #sTTAtPosMinus90Done )
   END_RUNG wire#w2
   RUNG wire#powerrail
      I_Contact( #iPos1Cmd )
      I_Contact( #iPos3Cmd )
      I_Contact( #iPos2Cmd )
      Contact( #iPos3StopSens )
   END_RUNG wire#w2
   // the same network as SCL:
   #qPos3Over := (#iPos3Cmd AND #iPos3StopSens AND (#sMinus90PosActiveForFwdOver OR #sMinus90PosActiveForRevOver OR #sTTAtPosMinus90Done)) OR (NOT #iPos1Cmd AND NOT #iPos3Cmd AND NOT #iPos2Cmd AND #iPos3StopSens);
END_REGION

REGION Network 18: Reset minus 90 forword and reverse command
   RUNG wire#powerrail
      Contact( #iPos3Cmd )
      Contact( #iPos3StopSens )
      wire#w1
      R_Coil( #sMinus90PosActiveForRev )
   END_RUNG
   RUNG wire#powerrail
      I_Contact( #iPos3Cmd )
   END_RUNG wire#w1
   // the same network as SCL:
   IF (#iPos3Cmd AND #iPos3StopSens) OR NOT #iPos3Cmd THEN #sMinus90PosActiveForRev := FALSE; END_IF;
END_REGION

REGION Network 19: Move to plus 90 degree
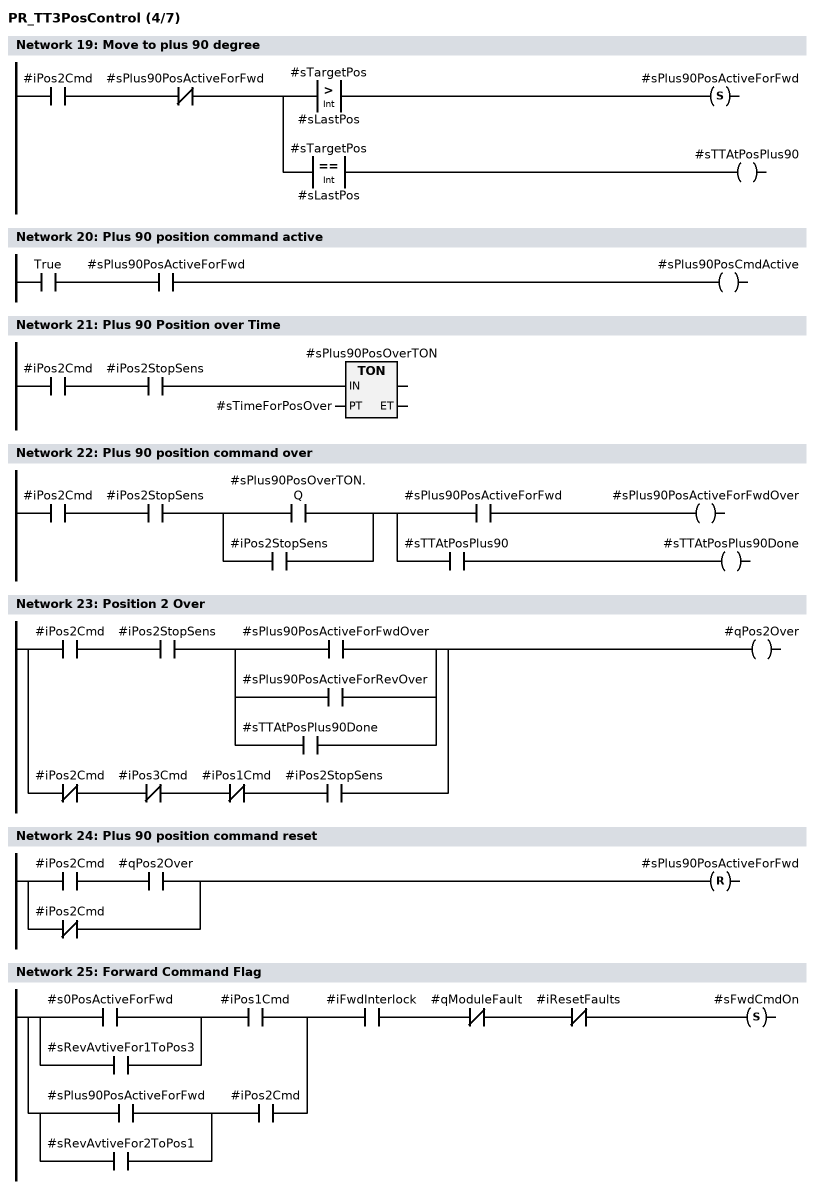
   RUNG wire#powerrail
      Contact( #iPos2Cmd )
      I_Contact( #sPlus90PosActiveForFwd )
      wire#w1
      { S7_Templates := "SrcType := Int" } GT_Contact(in1 := #sTargetPos, in2 := #sLastPos)
      S_Coil( #sPlus90PosActiveForFwd )
   END_RUNG
   RUNG wire#w1
      { S7_Templates := "SrcType := Int" } EQ_Contact(in1 := #sTargetPos, in2 := #sLastPos)
      Coil( #sTTAtPosPlus90 )
   END_RUNG
   // the same network as SCL:
   #_w1 := #iPos2Cmd AND NOT #sPlus90PosActiveForFwd;
   IF #_w1 AND (#sTargetPos > #sLastPos) THEN #sPlus90PosActiveForFwd := TRUE; END_IF;
   #sTTAtPosPlus90 := #_w1 AND (#sTargetPos = #sLastPos);
END_REGION

REGION Network 20: Plus 90 position command active
   RUNG wire#powerrail
      Contact( True )
      Contact( #sPlus90PosActiveForFwd )
      Coil( #sPlus90PosCmdActive )
   END_RUNG
   // the same network as SCL:
   #sPlus90PosCmdActive := True AND #sPlus90PosActiveForFwd;
END_REGION

REGION Network 21: Plus 90 Position over Time
   #sPlus90PosOverTON(IN := #iPos2Cmd AND #iPos2StopSens, PT := #sTimeForPosOver);   // TON
END_REGION

REGION Network 22: Plus 90 position command over
   RUNG wire#powerrail
      Contact( #iPos2Cmd )
      Contact( #iPos2StopSens )
      wire#w1
      Contact( #sPlus90PosOverTON.Q )
      wire#w2
      Contact( #sPlus90PosActiveForFwd )
      Coil( #sPlus90PosActiveForFwdOver )
   END_RUNG
   RUNG wire#w1
      Contact( #iPos2StopSens )
   END_RUNG wire#w2
   RUNG wire#w2
      Contact( #sTTAtPosPlus90 )
      Coil( #sTTAtPosPlus90Done )
   END_RUNG
   // the same network as SCL:
   #_w1 := #iPos2Cmd AND #iPos2StopSens AND (#sPlus90PosOverTON.Q OR #iPos2StopSens);
   #sPlus90PosActiveForFwdOver := #_w1 AND #sPlus90PosActiveForFwd;
   #sTTAtPosPlus90Done := #_w1 AND #sTTAtPosPlus90;
END_REGION

REGION Network 23: Position 2 Over
   RUNG wire#powerrail
      Contact( #iPos2Cmd )
      Contact( #iPos2StopSens )
      wire#w1
      Contact( #sPlus90PosActiveForFwdOver )
      wire#w2
      Coil( #qPos2Over )
   END_RUNG
   RUNG wire#w1
      Contact( #sPlus90PosActiveForRevOver )
   END_RUNG wire#w2
   RUNG wire#w1
      Contact( #sTTAtPosPlus90Done )
   END_RUNG wire#w2
   RUNG wire#powerrail
      I_Contact( #iPos2Cmd )
      I_Contact( #iPos3Cmd )
      I_Contact( #iPos1Cmd )
      Contact( #iPos2StopSens )
   END_RUNG wire#w2
   // the same network as SCL:
   #qPos2Over := (#iPos2Cmd AND #iPos2StopSens AND (#sPlus90PosActiveForFwdOver OR #sPlus90PosActiveForRevOver OR #sTTAtPosPlus90Done)) OR (NOT #iPos2Cmd AND NOT #iPos3Cmd AND NOT #iPos1Cmd AND #iPos2StopSens);
END_REGION

REGION Network 24: Plus 90 position command reset
   RUNG wire#powerrail
      Contact( #iPos2Cmd )
      Contact( #qPos2Over )
      wire#w1
      R_Coil( #sPlus90PosActiveForFwd )
   END_RUNG
   RUNG wire#powerrail
      I_Contact( #iPos2Cmd )
   END_RUNG wire#w1
   // the same network as SCL:
   IF (#iPos2Cmd AND #qPos2Over) OR NOT #iPos2Cmd THEN #sPlus90PosActiveForFwd := FALSE; END_IF;
END_REGION

REGION Network 25: Forward Command Flag
   RUNG wire#powerrail
      Contact( #s0PosActiveForFwd )
      wire#w1
      Contact( #iPos1Cmd )
      wire#w2
      Contact( #iFwdInterlock )
      I_Contact( #qModuleFault )
      I_Contact( #iResetFaults )
      S_Coil( #sFwdCmdOn )
   END_RUNG
   RUNG wire#powerrail
      Contact( #sRevAvtiveFor1ToPos3 )
   END_RUNG wire#w1
   RUNG wire#powerrail
      Contact( #sPlus90PosActiveForFwd )
      wire#w3
      Contact( #iPos2Cmd )
   END_RUNG wire#w2
   RUNG wire#powerrail
      Contact( #sRevAvtiveFor2ToPos1 )
   END_RUNG wire#w3
   // the same network as SCL:
   IF (((#s0PosActiveForFwd OR #sRevAvtiveFor1ToPos3) AND #iPos1Cmd) OR ((#sPlus90PosActiveForFwd OR #sRevAvtiveFor2ToPos1) AND #iPos2Cmd)) AND #iFwdInterlock AND NOT #qModuleFault AND NOT #iResetFaults THEN
       #sFwdCmdOn := TRUE;
   END_IF;
END_REGION

REGION Network 26: Reverse Command Flag
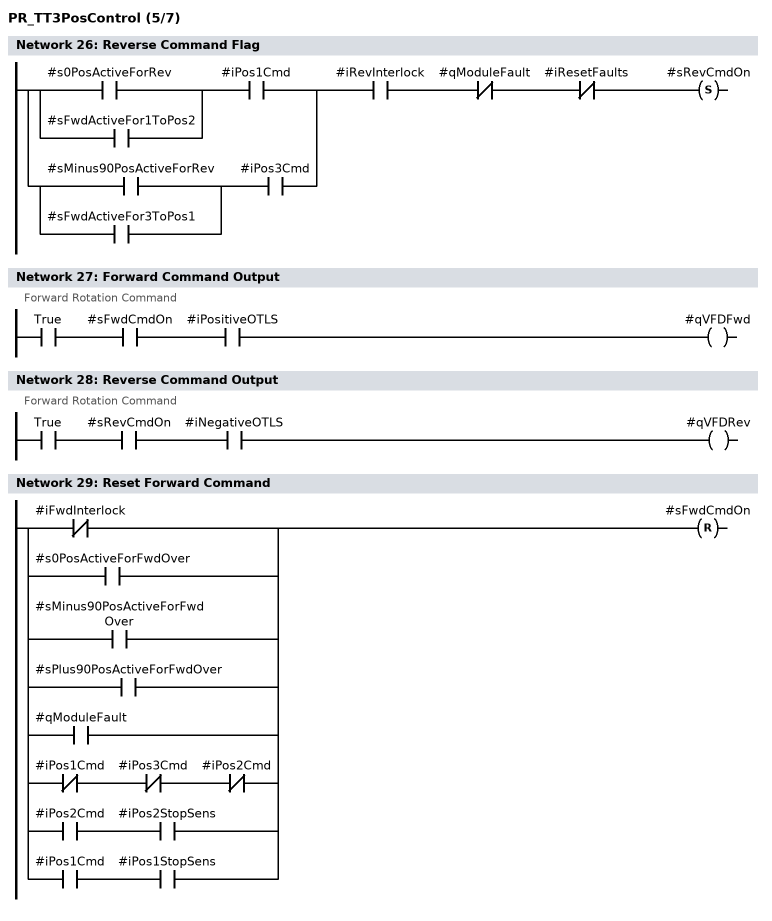
   RUNG wire#powerrail
      Contact( #s0PosActiveForRev )
      wire#w1
      Contact( #iPos1Cmd )
      wire#w2
      Contact( #iRevInterlock )
      I_Contact( #qModuleFault )
      I_Contact( #iResetFaults )
      S_Coil( #sRevCmdOn )
   END_RUNG
   RUNG wire#powerrail
      Contact( #sFwdActiveFor1ToPos2 )
   END_RUNG wire#w1
   RUNG wire#powerrail
      Contact( #sMinus90PosActiveForRev )
      wire#w3
      Contact( #iPos3Cmd )
   END_RUNG wire#w2
   RUNG wire#powerrail
      Contact( #sFwdActiveFor3ToPos1 )
   END_RUNG wire#w3
   // the same network as SCL:
   IF (((#s0PosActiveForRev OR #sFwdActiveFor1ToPos2) AND #iPos1Cmd) OR ((#sMinus90PosActiveForRev OR #sFwdActiveFor3ToPos1) AND #iPos3Cmd)) AND #iRevInterlock AND NOT #qModuleFault AND NOT #iResetFaults THEN
       #sRevCmdOn := TRUE;
   END_IF;
END_REGION

REGION Network 27: Forward Command Output
   // Forward Rotation Command
   RUNG wire#powerrail
      Contact( True )
      Contact( #sFwdCmdOn )
      Contact( #iPositiveOTLS )
      Coil( #qVFDFwd )
   END_RUNG
   // the same network as SCL:
   #qVFDFwd := True AND #sFwdCmdOn AND #iPositiveOTLS;
END_REGION

REGION Network 28: Reverse Command Output
   // Forward Rotation Command
   RUNG wire#powerrail
      Contact( True )
      Contact( #sRevCmdOn )
      Contact( #iNegativeOTLS )
      Coil( #qVFDRev )
   END_RUNG
   // the same network as SCL:
   #qVFDRev := True AND #sRevCmdOn AND #iNegativeOTLS;
END_REGION

REGION Network 29: Reset Forward Command
   RUNG wire#powerrail
      I_Contact( #iFwdInterlock )
      wire#w1
      R_Coil( #sFwdCmdOn )
   END_RUNG
   RUNG wire#powerrail
      Contact( #s0PosActiveForFwdOver )
   END_RUNG wire#w1
   RUNG wire#powerrail
      Contact( #sMinus90PosActiveForFwdOver )
   END_RUNG wire#w1
   RUNG wire#powerrail
      Contact( #sPlus90PosActiveForFwdOver )
   END_RUNG wire#w1
   RUNG wire#powerrail
      Contact( #qModuleFault )
   END_RUNG wire#w1
   RUNG wire#powerrail
      I_Contact( #iPos1Cmd )
      I_Contact( #iPos3Cmd )
      I_Contact( #iPos2Cmd )
   END_RUNG wire#w1
   RUNG wire#powerrail
      Contact( #iPos2Cmd )
      Contact( #iPos2StopSens )
   END_RUNG wire#w1
   RUNG wire#powerrail
      Contact( #iPos1Cmd )
      Contact( #iPos1StopSens )
   END_RUNG wire#w1
   // the same network as SCL:
   IF NOT #iFwdInterlock OR #s0PosActiveForFwdOver OR #sMinus90PosActiveForFwdOver OR #sPlus90PosActiveForFwdOver OR #qModuleFault OR (NOT #iPos1Cmd AND NOT #iPos3Cmd AND NOT #iPos2Cmd) OR (#iPos2Cmd AND #iPos2StopSens) OR (#iPos1Cmd AND #iPos1StopSens) THEN
       #sFwdCmdOn := FALSE;
   END_IF;
END_REGION

REGION Network 30: Reset Reverse Command
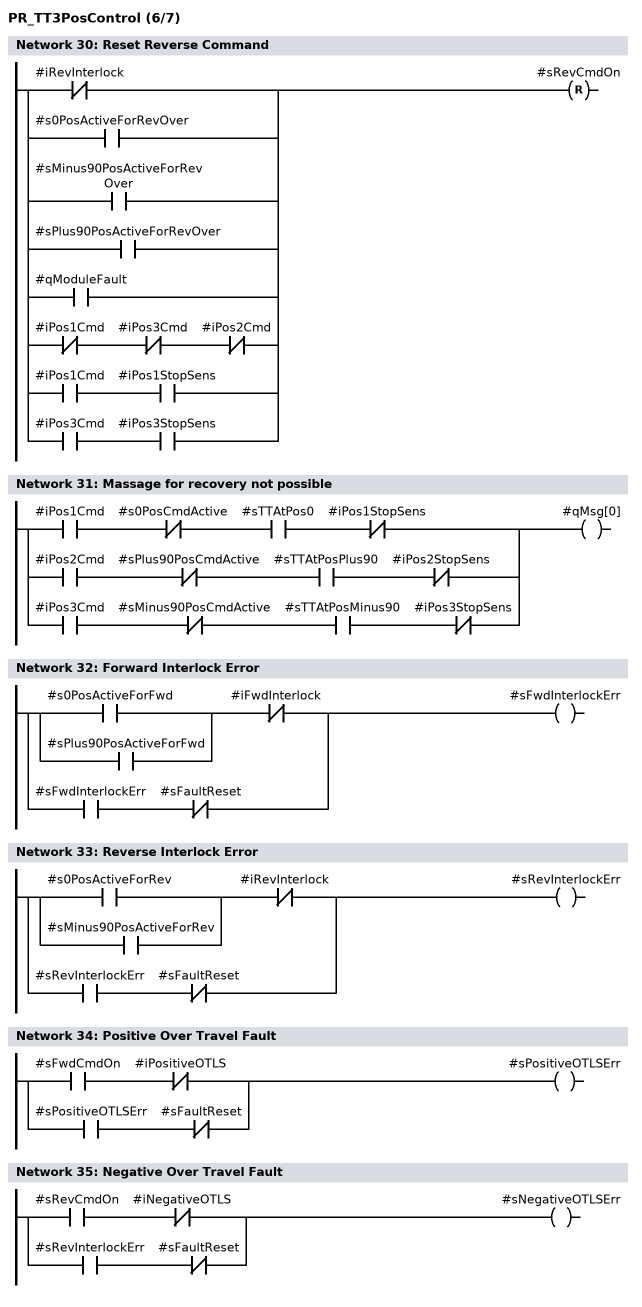
   RUNG wire#powerrail
      I_Contact( #iRevInterlock )
      wire#w1
      R_Coil( #sRevCmdOn )
   END_RUNG
   RUNG wire#powerrail
      Contact( #s0PosActiveForRevOver )
   END_RUNG wire#w1
   RUNG wire#powerrail
      Contact( #sMinus90PosActiveForRevOver )
   END_RUNG wire#w1
   RUNG wire#powerrail
      Contact( #sPlus90PosActiveForRevOver )
   END_RUNG wire#w1
   RUNG wire#powerrail
      Contact( #qModuleFault )
   END_RUNG wire#w1
   RUNG wire#powerrail
      I_Contact( #iPos1Cmd )
      I_Contact( #iPos3Cmd )
      I_Contact( #iPos2Cmd )
   END_RUNG wire#w1
   RUNG wire#powerrail
      Contact( #iPos1Cmd )
      Contact( #iPos1StopSens )
   END_RUNG wire#w1
   RUNG wire#powerrail
      Contact( #iPos3Cmd )
      Contact( #iPos3StopSens )
   END_RUNG wire#w1
   // the same network as SCL:
   IF NOT #iRevInterlock OR #s0PosActiveForRevOver OR #sMinus90PosActiveForRevOver OR #sPlus90PosActiveForRevOver OR #qModuleFault OR (NOT #iPos1Cmd AND NOT #iPos3Cmd AND NOT #iPos2Cmd) OR (#iPos1Cmd AND #iPos1StopSens) OR (#iPos3Cmd AND #iPos3StopSens) THEN
       #sRevCmdOn := FALSE;
   END_IF;
END_REGION

REGION Network 31: Massage for recovery not possible
   RUNG wire#powerrail
      Contact( #iPos1Cmd )
      I_Contact( #s0PosCmdActive )
      Contact( #sTTAtPos0 )
      I_Contact( #iPos1StopSens )
      wire#w1
      Coil( #qMsg[0] )
   END_RUNG
   RUNG wire#powerrail
      Contact( #iPos2Cmd )
      I_Contact( #sPlus90PosCmdActive )
      Contact( #sTTAtPosPlus90 )
      I_Contact( #iPos2StopSens )
   END_RUNG wire#w1
   RUNG wire#powerrail
      Contact( #iPos3Cmd )
      I_Contact( #sMinus90PosCmdActive )
      Contact( #sTTAtPosMinus90 )
      I_Contact( #iPos3StopSens )
   END_RUNG wire#w1
   // the same network as SCL:
   #qMsg[0] := (#iPos1Cmd AND NOT #s0PosCmdActive AND #sTTAtPos0 AND NOT #iPos1StopSens) OR (#iPos2Cmd AND NOT #sPlus90PosCmdActive AND #sTTAtPosPlus90 AND NOT #iPos2StopSens) OR (#iPos3Cmd AND NOT #sMinus90PosCmdActive AND #sTTAtPosMinus90 AND NOT #iPos3StopSens);
END_REGION

REGION Network 32: Forward Interlock Error
   RUNG wire#powerrail
      Contact( #s0PosActiveForFwd )
      wire#w1
      I_Contact( #iFwdInterlock )
      wire#w2
      Coil( #sFwdInterlockErr )
   END_RUNG
   RUNG wire#powerrail
      Contact( #sPlus90PosActiveForFwd )
   END_RUNG wire#w1
   RUNG wire#powerrail
      Contact( #sFwdInterlockErr )
      I_Contact( #sFaultReset )
   END_RUNG wire#w2
   // the same network as SCL:
   #sFwdInterlockErr := ((#s0PosActiveForFwd OR #sPlus90PosActiveForFwd) AND NOT #iFwdInterlock) OR (#sFwdInterlockErr AND NOT #sFaultReset);
END_REGION

REGION Network 33: Reverse Interlock Error
   RUNG wire#powerrail
      Contact( #s0PosActiveForRev )
      wire#w1
      I_Contact( #iRevInterlock )
      wire#w2
      Coil( #sRevInterlockErr )
   END_RUNG
   RUNG wire#powerrail
      Contact( #sMinus90PosActiveForRev )
   END_RUNG wire#w1
   RUNG wire#powerrail
      Contact( #sRevInterlockErr )
      I_Contact( #sFaultReset )
   END_RUNG wire#w2
   // the same network as SCL:
   #sRevInterlockErr := ((#s0PosActiveForRev OR #sMinus90PosActiveForRev) AND NOT #iRevInterlock) OR (#sRevInterlockErr AND NOT #sFaultReset);
END_REGION

REGION Network 34: Positive Over Travel Fault
   RUNG wire#powerrail
      Contact( #sFwdCmdOn )
      I_Contact( #iPositiveOTLS )
      wire#w1
      Coil( #sPositiveOTLSErr )
   END_RUNG
   RUNG wire#powerrail
      Contact( #sPositiveOTLSErr )
      I_Contact( #sFaultReset )
   END_RUNG wire#w1
   // the same network as SCL:
   #sPositiveOTLSErr := (#sFwdCmdOn AND NOT #iPositiveOTLS) OR (#sPositiveOTLSErr AND NOT #sFaultReset);
END_REGION

REGION Network 35: Negative Over Travel Fault
   RUNG wire#powerrail
      Contact( #sRevCmdOn )
      I_Contact( #iNegativeOTLS )
      wire#w1
      Coil( #sNegativeOTLSErr )
   END_RUNG
   RUNG wire#powerrail
      Contact( #sRevInterlockErr )
      I_Contact( #sFaultReset )
   END_RUNG wire#w1
   // the same network as SCL:
   #sNegativeOTLSErr := (#sRevCmdOn AND NOT #iNegativeOTLS) OR (#sRevInterlockErr AND NOT #sFaultReset);
END_REGION

REGION Network 36: Time out value validation for VFD stop
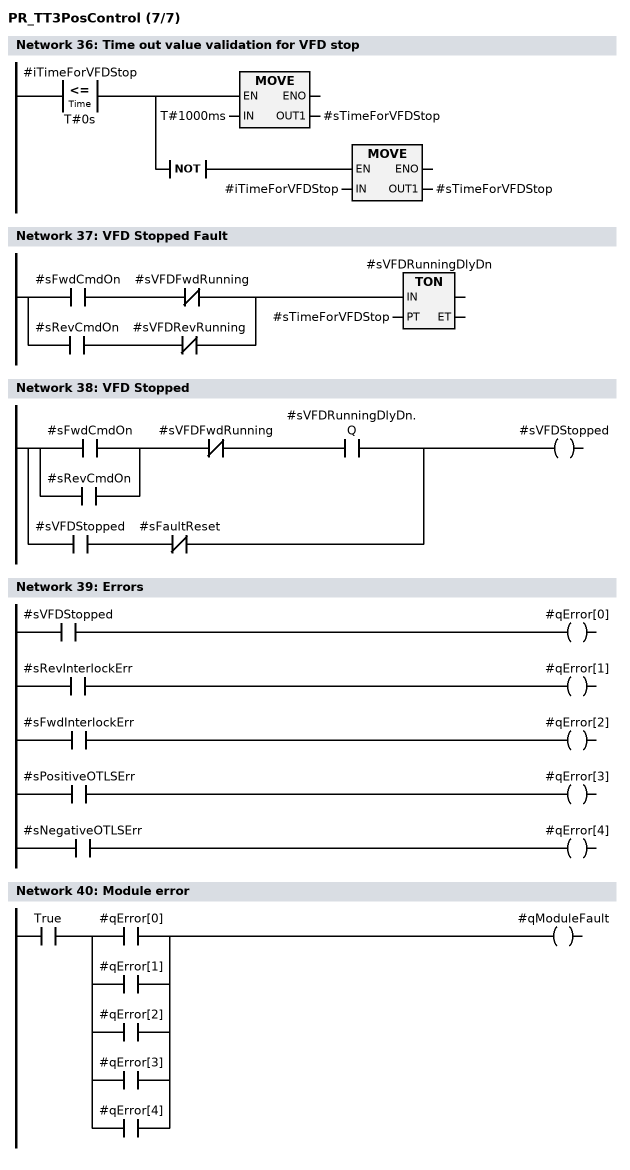
   RUNG wire#powerrail
      { S7_Templates := "SrcType := Time" } LE_Contact(in1 := #iTimeForVFDStop, in2 := T#0s)
      wire#w1
      Move(in := T#1000ms, out1 => #sTimeForVFDStop)
   END_RUNG
   RUNG wire#w1
      Not()
      Move(in := #iTimeForVFDStop, out1 => #sTimeForVFDStop)
   END_RUNG
   // the same network as SCL:
   #_w1 := #iTimeForVFDStop <= T#0s;
   IF #_w1 THEN #sTimeForVFDStop := T#1000ms; END_IF;
   IF NOT #_w1 THEN #sTimeForVFDStop := #iTimeForVFDStop; END_IF;
END_REGION

REGION Network 37: VFD Stopped Fault
   #sVFDRunningDlyDn(IN := (#sFwdCmdOn AND NOT #sVFDFwdRunning) OR (#sRevCmdOn AND NOT #sVFDRevRunning),   // TON
                     PT := #sTimeForVFDStop);
END_REGION

REGION Network 38: VFD Stopped
   RUNG wire#powerrail
      Contact( #sFwdCmdOn )
      wire#w1
      I_Contact( #sVFDFwdRunning )
      Contact( #sVFDRunningDlyDn.Q )
      wire#w2
      Coil( #sVFDStopped )
   END_RUNG
   RUNG wire#powerrail
      Contact( #sRevCmdOn )
   END_RUNG wire#w1
   RUNG wire#powerrail
      Contact( #sVFDStopped )
      I_Contact( #sFaultReset )
   END_RUNG wire#w2
   // the same network as SCL:
   #sVFDStopped := ((#sFwdCmdOn OR #sRevCmdOn) AND NOT #sVFDFwdRunning AND #sVFDRunningDlyDn.Q) OR (#sVFDStopped AND NOT #sFaultReset);
END_REGION

REGION Network 39: Errors
   RUNG wire#powerrail
      Contact( #sVFDStopped )
      Coil( #qError[0] )
   END_RUNG
   RUNG wire#powerrail
      Contact( #sRevInterlockErr )
      Coil( #qError[1] )
   END_RUNG
   RUNG wire#powerrail
      Contact( #sFwdInterlockErr )
      Coil( #qError[2] )
   END_RUNG
   RUNG wire#powerrail
      Contact( #sPositiveOTLSErr )
      Coil( #qError[3] )
   END_RUNG
   RUNG wire#powerrail
      Contact( #sNegativeOTLSErr )
      Coil( #qError[4] )
   END_RUNG
   // the same network as SCL:
   #qError[0] := #sVFDStopped;
   #qError[1] := #sRevInterlockErr;
   #qError[2] := #sFwdInterlockErr;
   #qError[3] := #sPositiveOTLSErr;
   #qError[4] := #sNegativeOTLSErr;
END_REGION

REGION Network 40: Module error
   RUNG wire#powerrail
      Contact( True )
      wire#w1
      Contact( #qError[0] )
      wire#w2
      Coil( #qModuleFault )
   END_RUNG
   RUNG wire#w1
      Contact( #qError[1] )
   END_RUNG wire#w2
   RUNG wire#w1
      Contact( #qError[2] )
   END_RUNG wire#w2
   RUNG wire#w1
      Contact( #qError[3] )
   END_RUNG wire#w2
   RUNG wire#w1
      Contact( #qError[4] )
   END_RUNG wire#w2
   // the same network as SCL:
   #qModuleFault := True AND (#qError[0] OR #qError[1] OR #qError[2] OR #qError[3] OR #qError[4]);
END_REGION
END_FUNCTION_BLOCK